(* IEC 61131-3 sources: TetherPLC/tests/fbd_gallery, 10 files *)

(* ---- 01_ton_debounce.st ---- *)
PROGRAM P01_TON_DEBOUNCE
VAR
    start_in AT %IX0.0 : BOOL;
    stop_in AT %IX0.1 : BOOL;
    run AT %QX0.0 : BOOL;
    ton1 : TON;
END_VAR
ton1(IN := start_in, PT := T#200ms);
run := ton1.Q AND NOT stop_in;
END_PROGRAM

(* ---- 02_ctu_count.st ---- *)
PROGRAM P02_CTU_COUNT
VAR
    pulse AT %IX0.0 : BOOL;
    reset AT %IX0.1 : BOOL;
    done AT %QX0.0 : BOOL;
    ctu1 : CTU;
END_VAR
ctu1(CU := pulse, R := reset, PV := 3);
done := ctu1.QU;
END_PROGRAM

(* ---- 03_sel_gate.st ---- *)
PROGRAM P03_SEL_GATE
VAR
    g AT %IX0.0 : BOOL;
    a AT %IB1 : BYTE;
    b AT %IB2 : BYTE;
    out AT %QB0 : BYTE;
END_VAR
IF g THEN
    out := b;
ELSE
    out := a;
END_IF;
END_PROGRAM

(* ---- 04_limit_clamp.st ---- *)
PROGRAM P04_LIMIT_CLAMP
VAR
    x AT %IB1 : BYTE;
    out AT %QB0 : BYTE;
END_VAR
IF x < 10 THEN
    out := 10;
ELSIF x > 200 THEN
    out := 200;
ELSE
    out := x;
END_IF;
END_PROGRAM

(* ---- 05_mux_pick.st ---- *)
PROGRAM P05_MUX_PICK
VAR
    k AT %IB1 : BYTE;
    out AT %QB0 : BYTE;
END_VAR
CASE k OF
    0: out := 10;
    1: out := 20;
    2: out := 30;
ELSE
    out := 10;
END_CASE;
END_PROGRAM

(* ---- 06_sr_latch.st ---- *)
PROGRAM P06_SR_LATCH
VAR
    s AT %IX0.0 : BOOL;
    r AT %IX0.1 : BOOL;
    q AT %QX0.0 : BOOL;
    sr1 : SR;
END_VAR
sr1(S1 := s, R := r);
q := sr1.Q1;
END_PROGRAM

(* ---- 07_two_nets.st ---- *)
PROGRAM P07_TWO_NETS
VAR
    a AT %IX0.0 : BOOL;
    b AT %IX0.1 : BOOL;
    q AT %QX0.0 : BOOL;
    gate : BOOL;
END_VAR
gate := a AND b;
q := gate;
END_PROGRAM

(* ---- 08_assoc_bind.st ---- *)
PROGRAM P08_ASSOC_BIND
VAR
    en_in AT %IX0.0 : BOOL;
    q AT %QX0.0 : BOOL;
END_VAR
q := en_in;
END_PROGRAM

(* ---- 09_cmp_ge.st ---- *)
PROGRAM P09_CMP_GE
VAR
    x AT %IB1 : BYTE;
    q AT %QX0.0 : BOOL;
END_VAR
q := x >= 100;
END_PROGRAM

(* ---- 10_tof_hold.st ---- *)
PROGRAM P10_TOF_HOLD
VAR
    x AT %IX0.0 : BOOL;
    q AT %QX0.0 : BOOL;
    tof1 : TOF;
END_VAR
tof1(IN := x, PT := T#200ms);
q := tof1.Q;
END_PROGRAM
